(* PLC project v0.5.3_PreCommissioningPrep.project, CODESYS CODESYS V3.5 SP19 Patch 1 *)
(* stored: creationDateTime 2026-07-29T10:07:35.239406, modificationDateTime 2026-07-28T11:53:41.5518987 *)

PROGRAM PRG_12_LD

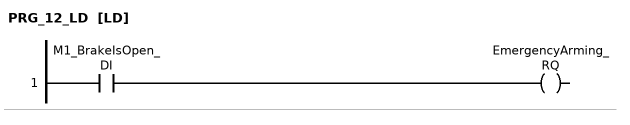
(* LD diagram, written out as Structured Text *)

EmergencyArming_RQ := M1_BrakeIsOpen_DI;
END_PROGRAM
